Fanuc KAREL source: KD00024.KL

PROGRAM KD00024
%NOLOCKGROUP
VAR
  I: INTEGER
  J: INTEGER
  B: BOOLEAN
  R: REAL
  S: STRING[80]
BEGIN
  I = 1
  CONDITION[1]:
  WHEN I > EVAL(10 * I) DO
    J = 1
  ENDCONDITION
END KD00024
